Universal Robots URScript: 1Johnathan.script

def output_0001():
  # Default parameters:
  global speed_ms = 0.3
  global speed_rads = 0.75
  global accel_mss = 3
  global accel_radss = 1.2
  global blend_radius_m = 0.001

  # Add subprograms here
  # Start of main program
  # Program generated by RoboDK v5.7.4 for UR10e on 22/07/2024 10:59:04
  # Using nominal kinematics.
  blend_radius_m = 0.001
  speed_ms = 1.000
  # set_reference(p[-0.375000, 0.265000, -0.018000, 0.000000, 0.000000, 0.000000])
  set_tcp(p[0.000000, 0.000000, 0.252000, 0.000000, 0.000000, 0.000000])
  # Show Tool
  movej([2.604293, -1.437179, -2.485600, -0.789610, 1.570796, -2.108096],accel_radss,speed_rads,0,blend_radius_m)
  movel([2.604293, -1.497217, -2.512761, -0.702411, 1.570796, -2.108096],accel_mss,speed_ms,0,blend_radius_m)
  speed_ms = 1.000
  speed_ms = 0.002
  movel([2.604293, -1.508175, -2.517063, -0.687151, 1.570796, -2.108096],accel_mss,speed_ms,0,blend_radius_m)
  speed_ms = 0.007
  movec([2.603816, -1.508462, -2.516806, -0.687120, 1.570796, -2.108573],[2.603307, -1.508637, -2.516650, -0.687102, 1.570796, -2.109082],accel_mss,speed_ms,blend_radius_m)
  movec([2.602757, -1.508696, -2.516598, -0.687096, 1.570796, -2.109632],[2.602268, -1.508621, -2.516664, -0.687104, 1.570796, -2.110121],accel_mss,speed_ms,blend_radius_m)
  movec([2.600447, -1.508284, -2.516966, -0.687139, 1.570796, -2.111942],[2.598423, -1.508336, -2.516919, -0.687134, 1.570796, -2.113966],accel_mss,speed_ms,blend_radius_m)
  movec([2.595446, -1.508878, -2.516434, -0.687077, 1.570796, -2.116943],[2.592433, -1.509794, -2.515613, -0.686982, 1.570796, -2.119956],accel_mss,speed_ms,blend_radius_m)
  movec([2.591318, -1.510221, -2.515230, -0.686938, 1.570796, -2.121071],[2.590209, -1.510687, -2.514812, -0.686890, 1.570796, -2.122180],accel_mss,speed_ms,blend_radius_m)
  movec([2.583631, -1.513609, -2.512179, -0.686601, 1.570796, -2.128758],[2.577095, -1.516580, -2.509488, -0.686321, 1.570796, -2.135294],accel_mss,speed_ms,blend_radius_m)
  movec([2.550168, -1.529181, -2.497909, -0.685299, 1.570796, -2.162221],[2.523831, -1.541945, -2.485907, -0.684537, 1.570796, -2.188558],accel_mss,speed_ms,blend_radius_m)
  movec([2.518527, -1.544567, -2.483408, -0.684414, 1.570796, -2.193862],[2.513247, -1.547191, -2.480895, -0.684304, 1.570796, -2.199142],accel_mss,speed_ms,blend_radius_m)
  movel([2.510802, -1.548411, -2.479722, -0.684256, 1.570796, -2.201587],accel_mss,speed_ms,0,blend_radius_m)
  movel([2.510282, -1.547905, -2.480209, -0.684275, 1.570796, -2.202107],accel_mss,speed_ms,0,blend_radius_m)
  movel([2.509762, -1.547398, -2.480695, -0.684295, 1.570796, -2.202627],accel_mss,speed_ms,0,blend_radius_m)
  movel([2.519376, -1.532909, -2.494432, -0.685048, 1.570796, -2.193013],accel_mss,speed_ms,0,blend_radius_m)
  movec([2.526773, -1.521882, -2.504648, -0.685858, 1.570796, -2.185616],[2.534360, -1.510676, -2.514822, -0.686891, 1.570796, -2.178029],accel_mss,speed_ms,blend_radius_m)
  movec([2.540243, -1.502051, -2.522508, -0.687830, 1.570796, -2.172146],[2.546242, -1.493314, -2.530168, -0.688907, 1.570796, -2.166147],accel_mss,speed_ms,blend_radius_m)
  movec([2.552500, -1.484076, -2.538129, -0.690184, 1.570796, -2.159889],[2.558671, -1.474659, -2.546100, -0.691631, 1.570796, -2.153718],accel_mss,speed_ms,blend_radius_m)
  movec([2.559369, -1.473377, -2.547173, -0.691839, 1.570796, -2.153020],[2.559821, -1.472092, -2.548247, -0.692050, 1.570796, -2.152568],accel_mss,speed_ms,blend_radius_m)
  movec([2.560032, -1.470863, -2.549271, -0.692255, 1.570796, -2.152357],[2.560031, -1.469688, -2.550248, -0.692453, 1.570796, -2.152358],accel_mss,speed_ms,blend_radius_m)
  movec([2.559843, -1.468863, -2.550933, -0.692594, 1.570796, -2.152546],[2.559447, -1.468147, -2.551525, -0.692716, 1.570796, -2.152941],accel_mss,speed_ms,blend_radius_m)
  movel([2.559402, -1.467478, -2.552079, -0.692832, 1.570796, -2.152987],accel_mss,speed_ms,0,blend_radius_m)
  movec([2.559662, -1.467023, -2.552455, -0.692911, 1.570796, -2.152727],[2.560056, -1.466607, -2.552799, -0.692983, 1.570796, -2.152333],accel_mss,speed_ms,blend_radius_m)
  movel([2.561141, -1.465689, -2.553556, -0.693144, 1.570796, -2.151248],accel_mss,speed_ms,0,blend_radius_m)
  movel([2.569602, -1.473225, -2.547300, -0.691864, 1.570796, -2.142787],accel_mss,speed_ms,0,blend_radius_m)
  movel([2.577874, -1.480796, -2.540921, -0.690671, 1.570796, -2.134515],accel_mss,speed_ms,0,blend_radius_m)
  movel([2.576802, -1.481675, -2.540175, -0.690539, 1.570796, -2.135587],accel_mss,speed_ms,0,blend_radius_m)
  movel([2.575732, -1.482552, -2.539429, -0.690408, 1.570796, -2.136657],accel_mss,speed_ms,0,blend_radius_m)
  movel([2.574373, -1.481546, -2.540285, -0.690558, 1.570796, -2.138016],accel_mss,speed_ms,0,blend_radius_m)
  movec([2.572968, -1.480689, -2.541012, -0.690687, 1.570796, -2.139420],[2.571366, -1.480046, -2.541558, -0.690785, 1.570796, -2.141023],accel_mss,speed_ms,blend_radius_m)
  movec([2.570473, -1.479905, -2.541678, -0.690807, 1.570796, -2.141916],[2.569470, -1.479998, -2.541598, -0.690792, 1.570796, -2.142919],accel_mss,speed_ms,blend_radius_m)
  movec([2.568854, -1.480172, -2.541451, -0.690766, 1.570796, -2.143535],[2.568245, -1.480441, -2.541223, -0.690725, 1.570796, -2.144144],accel_mss,speed_ms,blend_radius_m)
  movec([2.567531, -1.480864, -2.540864, -0.690661, 1.570796, -2.144858],[2.566868, -1.481359, -2.540443, -0.690586, 1.570796, -2.145521],accel_mss,speed_ms,blend_radius_m)
  movec([2.565928, -1.482228, -2.539705, -0.690456, 1.570796, -2.146461],[2.565112, -1.483163, -2.538908, -0.690318, 1.570796, -2.147277],accel_mss,speed_ms,blend_radius_m)
  movec([2.560639, -1.489029, -2.533878, -0.689482, 1.570796, -2.151750],[2.556366, -1.494884, -2.528801, -0.688704, 1.570796, -2.156023],accel_mss,speed_ms,blend_radius_m)
  movel([2.549296, -1.504827, -2.520047, -0.687514, 1.570796, -2.163093],accel_mss,speed_ms,0,blend_radius_m)
  movel([2.557748, -1.512187, -2.513462, -0.686740, 1.570796, -2.154641],accel_mss,speed_ms,0,blend_radius_m)
  movel([2.566016, -1.519585, -2.506751, -0.686053, 1.570796, -2.146373],accel_mss,speed_ms,0,blend_radius_m)
  movel([2.567160, -1.519061, -2.507230, -0.686099, 1.570796, -2.145229],accel_mss,speed_ms,0,blend_radius_m)
  movec([2.573813, -1.515998, -2.510017, -0.686374, 1.570796, -2.138576],[2.580487, -1.512895, -2.512824, -0.686670, 1.570796, -2.131902],accel_mss,speed_ms,blend_radius_m)
  movec([2.582441, -1.511953, -2.513673, -0.686763, 1.570796, -2.129948],[2.584381, -1.510962, -2.514565, -0.686862, 1.570796, -2.128008],accel_mss,speed_ms,blend_radius_m)
  movec([2.588316, -1.508472, -2.516798, -0.687119, 1.570796, -2.124073],[2.591759, -1.505418, -2.519523, -0.687449, 1.570796, -2.120630],accel_mss,speed_ms,blend_radius_m)
  movec([2.593122, -1.503401, -2.521314, -0.687675, 1.570796, -2.119267],[2.593472, -1.501385, -2.523097, -0.687908, 1.570796, -2.118917],accel_mss,speed_ms,blend_radius_m)
  movec([2.593279, -1.500404, -2.523962, -0.688023, 1.570796, -2.119110],[2.592918, -1.499503, -2.524755, -0.688131, 1.570796, -2.119471],accel_mss,speed_ms,blend_radius_m)
  movec([2.592299, -1.498508, -2.525630, -0.688251, 1.570796, -2.120090],[2.591523, -1.497619, -2.526410, -0.688360, 1.570796, -2.120866],accel_mss,speed_ms,blend_radius_m)
  movec([2.591147, -1.497231, -2.526749, -0.688408, 1.570796, -2.121242],[2.590794, -1.496826, -2.527104, -0.688459, 1.570796, -2.121595],accel_mss,speed_ms,blend_radius_m)
  movel([2.590775, -1.496714, -2.527203, -0.688473, 1.570796, -2.121614],accel_mss,speed_ms,0,blend_radius_m)
  movel([2.590862, -1.496591, -2.527310, -0.688488, 1.570796, -2.121527],accel_mss,speed_ms,0,blend_radius_m)
  movec([2.591353, -1.496203, -2.527649, -0.688537, 1.570796, -2.121036],[2.591858, -1.495830, -2.527975, -0.688584, 1.570796, -2.120531],accel_mss,speed_ms,blend_radius_m)
  movel([2.592904, -1.495083, -2.528627, -0.688679, 1.570796, -2.119485],accel_mss,speed_ms,0,blend_radius_m)
  movel([2.599163, -1.501241, -2.523224, -0.687924, 1.570796, -2.113226],accel_mss,speed_ms,0,blend_radius_m)
  movel([2.605310, -1.507412, -2.517745, -0.687232, 1.570796, -2.107079],accel_mss,speed_ms,0,blend_radius_m)
  movel([2.604293, -1.508175, -2.517063, -0.687151, 1.570796, -2.108096],accel_mss,speed_ms,0,blend_radius_m)
  speed_ms = 1.000
  movel([2.604293, -1.497217, -2.512761, -0.702411, 1.570796, -2.108096],accel_mss,speed_ms,0,blend_radius_m)
  movel([2.547578, -1.496299, -2.513567, -0.702524, 1.570796, -2.164811],accel_mss,speed_ms,0,blend_radius_m)
  speed_ms = 0.002
  movel([2.547578, -1.507268, -2.517873, -0.687247, 1.570796, -2.164811],accel_mss,speed_ms,0,blend_radius_m)
  speed_ms = 0.007
  movec([2.536165, -1.522961, -2.503658, -0.685770, 1.570796, -2.176224],[2.525389, -1.538371, -2.489295, -0.684723, 1.570796, -2.187000],accel_mss,speed_ms,blend_radius_m)
  movec([2.525242, -1.538815, -2.488876, -0.684698, 1.570796, -2.187147],[2.525421, -1.539153, -2.488556, -0.684680, 1.570796, -2.186968],accel_mss,speed_ms,blend_radius_m)
  movec([2.525785, -1.539248, -2.488466, -0.684675, 1.570796, -2.186604],[2.526231, -1.539131, -2.488577, -0.684681, 1.570796, -2.186157],accel_mss,speed_ms,blend_radius_m)
  movec([2.544519, -1.530130, -2.497026, -0.685233, 1.570796, -2.167870],[2.563046, -1.521033, -2.505427, -0.685929, 1.570796, -2.149343],accel_mss,speed_ms,blend_radius_m)
  movel([2.563102, -1.520908, -2.505541, -0.685940, 1.570796, -2.149287],accel_mss,speed_ms,0,blend_radius_m)
  movec([2.559485, -1.517496, -2.508655, -0.686238, 1.570796, -2.152904],[2.555780, -1.514131, -2.511708, -0.686550, 1.570796, -2.156609],accel_mss,speed_ms,blend_radius_m)
  movec([2.551967, -1.510750, -2.514755, -0.686884, 1.570796, -2.160422],[2.548119, -1.507375, -2.517779, -0.687236, 1.570796, -2.164270],accel_mss,speed_ms,blend_radius_m)
  movel([2.547936, -1.507201, -2.517934, -0.687255, 1.570796, -2.164453],accel_mss,speed_ms,0,blend_radius_m)
  movel([2.547751, -1.507159, -2.517971, -0.687259, 1.570796, -2.164638],accel_mss,speed_ms,0,blend_radius_m)
  movel([2.547578, -1.507268, -2.517873, -0.687247, 1.570796, -2.164811],accel_mss,speed_ms,0,blend_radius_m)
  speed_ms = 1.000
  movel([2.547578, -1.496299, -2.513567, -0.702524, 1.570796, -2.164811],accel_mss,speed_ms,0,blend_radius_m)
  movel([2.915402, -1.462227, -2.542486, -0.707676, 1.570796, -1.796986],accel_mss,speed_ms,0,blend_radius_m)
  movel([2.915402, -1.400124, -2.514210, -0.798055, 1.570796, -1.796986],accel_mss,speed_ms,0,blend_radius_m)
  # End of main program
end

output_0001()
